// =============================================================================
// s7-to-codesys — корпус SCL. Написан с нуля, объект вымышленный (ВОС «Северная»).
//
// Файл:   FB_BatchCounter.scl
// Блок:   FUNCTION_BLOCK "FB_BatchCounter"
// -----------------------------------------------------------------------------
// Назначение
//   Счёт доз реагента: импульсный расходомер дозирующего насоса даёт импульс
//   на каждые 10 мл; pulsesPerDose импульсов — одна доза; batchPreset доз —
//   партия (сигнал на смену бака). Экземпляр DB_Dosing.
//
// Логика (нормативное описание)
//   1. Импульс считается по спаду pulseInput (F_TRIG; контакт геркона
//      нормально замкнутый). reset (уровень) обнуляет счёт импульсов и счётчик доз.
//   2. pulseCounter := pulseCounter + 1 на каждый импульс; при
//      pulseCounter >= pulsesPerDose: doseDone (импульс на вызов) := TRUE,
//      pulseCounter := 0.
//   3. Счётчик доз — CTU_INT (CU := doseDone, R := reset, PV := batchPreset):
//      doseCount := CV, batchDone := Q.
//   4. statusByte: бит 0 — batchDone, бит 1 — счёт идёт (pulseCounter > 0),
//      бит 2 — pulsesPerDose <= 0 (ошибка параметра), биты 3...7 = 0.
//   5. packedCounters (DWord): старшее слово — doseCount, младшее — pulseCounter
//      (SHL на 16 и OR). lowWordCopy := packedCounters.%W0 (младшее слово),
//      highByteOfLow := lowWordCopy.%B1 (обращение к срезам).
// Что проверяет при конвертации
//   CTU_INT (в CODESYS у CTU вход RESET и тип WORD — нужна проверка), F_TRIG,
//   Byte/Word/DWord, SHL, OR, INT_TO_WORD, WORD_TO_DWORD, срезы .%Xn/.%Wn/.%Bn.
// =============================================================================
FUNCTION_BLOCK "FB_BatchCounter"
TITLE = Dosing pulse and batch counter
{ S7_Optimized_Access := 'TRUE' }
AUTHOR : WTP2
FAMILY : Dosing
VERSION : 1.1
   VAR_INPUT
      pulseInput : Bool;   // Импульсы расходомера реагента (НЗ контакт)
      reset : Bool;   // Сброс счёта (уровень)
      pulsesPerDose : Int := 100;   // Импульсов на одну дозу
      batchPreset : Int := 20;   // Доз в партии
   END_VAR

   VAR_OUTPUT
      doseDone : Bool;   // Доза набрана (один вызов)
      doseCount : Int;   // Число доз в партии
      batchDone : Bool;   // Партия набрана
      statusByte : Byte;   // Состояние для HMI
      packedCounters : DWord;   // Счётчики одним словом для верхнего уровня
      lowWordCopy : Word;   // Младшее слово packedCounters
      highByteOfLow : Byte;   // Старший байт младшего слова
   END_VAR

   VAR
      pulseCounter : Int;   // Импульсы текущей дозы
      edgePulse {InstructionName := 'F_TRIG'; LibVersion := '1.0'} : F_TRIG;
      ctuBatch {InstructionName := 'CTU_INT'; LibVersion := '1.0'} : CTU_INT;
   END_VAR


BEGIN
    REGION Pulses
        #edgePulse(CLK := #pulseInput);
        #doseDone := FALSE;
        IF #reset THEN
            #pulseCounter := 0;
        ELSIF #edgePulse.Q THEN
            #pulseCounter := #pulseCounter + 1;
            IF #pulsesPerDose > 0 AND #pulseCounter >= #pulsesPerDose THEN
                #doseDone := TRUE;
                #pulseCounter := 0;
            END_IF;
        END_IF;
    END_REGION

    REGION Batch counter
        #ctuBatch(CU := #doseDone,
                  R := #reset,
                  PV := #batchPreset);
        #doseCount := #ctuBatch.CV;
        #batchDone := #ctuBatch.Q;
    END_REGION

    REGION Status and packing
        #statusByte := 16#00;
        #statusByte.%X0 := #batchDone;
        #statusByte.%X1 := #pulseCounter > 0;
        #statusByte.%X2 := #pulsesPerDose <= 0;

        #packedCounters := SHL(IN := WORD_TO_DWORD(INT_TO_WORD(#doseCount)), N := 16)
                           OR WORD_TO_DWORD(INT_TO_WORD(#pulseCounter));
        #lowWordCopy := #packedCounters.%W0;
        #highByteOfLow := #lowWordCopy.%B1;
    END_REGION

END_FUNCTION_BLOCK

